// TIA Portal V20 export
FUNCTION_BLOCK "POS3_0_SK_Ablauf"   // FB26, GRAPH
// stored: GraphVersion 6.0, InitialValuesAcquisition false, LanguageInNetworks FBD, SetENOAutomatically false
   // inherited from GRAPH_BASE
   VAR_INPUT
      OFF_SQ { ExternalWritable := 'False'} : Bool := false;   // Kette ausschalten
      INIT_SQ { ExternalWritable := 'False'} : Bool := false;   // Kette in Initialzustand versetzen
      ACK_EF { ExternalWritable := 'False'} : Bool := false;   // Alle Fehler und Störungen quittieren
      REG_EF { ExternalWritable := 'False'} : Bool := false;   // Alle Fehler und Störungen registrieren
      ACK_S { ExternalWritable := 'False'} : Bool := false;   // Schritt quittieren, der an Parameter S_NO anliegt
      REG_S { ExternalWritable := 'False'} : Bool := false;   // Schritt registrieren, der an Parameter S_NO anliegt
      HALT_SQ { ExternalWritable := 'False'} : Bool := false;   // Kette sofort anhalten
      HALT_TM { ExternalWritable := 'False'} : Bool := false;   // Zeiten sofort anhalten
      ZERO_OP { ExternalWritable := 'False'} : Bool := false;   // Alle mit N, L, D zugewiesenen Operanden auf 0 setzen
      EN_IL { ExternalWritable := 'False'} : Bool := false;   // Interlockbearbeitung aktivieren
      EN_SV { ExternalWritable := 'False'} : Bool := false;   // Supervisionsbearbeitung aktivieren
      EN_ACKREQ { ExternalWritable := 'False'} : Bool := false;   // Quittierpflicht aktivieren
      EN_SSKIP { ExternalWritable := 'False'} : Bool := false;   // "Schritte überspringen" aktivieren
      DISP_SACT { ExternalWritable := 'False'} : Bool := false;   // Nur aktive Schritte anzeigen
      DISP_SEF { ExternalWritable := 'False'} : Bool := false;   // Nur fehlerhafte und gestörte Schritte anzeigen
      DISP_SALL { ExternalWritable := 'False'} : Bool := false;   // Alle Schritte anzeigen
      S_PREV { ExternalWritable := 'False'} : Bool := false;   // Vorherigen Schritt am Parameter S_NO ausgeben
      S_NEXT { ExternalWritable := 'False'} : Bool := false;   // Nächsten Schritt am Parameter S_NO anzeigen
      SW_AUTO { ExternalWritable := 'False'} : Bool := false;   // Automatischer Betrieb
      SW_TAP { ExternalWritable := 'False'} : Bool := false;   // Halbautomatisch/Weiterschalten mit Transition
      SW_TOP { ExternalWritable := 'False'} : Bool := false;   // Halbautomatisch/Ignoriere Transition
      SW_MAN { ExternalWritable := 'False'} : Bool := false;   // Handbetrieb
      S_SEL { ExternalWritable := 'False'} : Int := 0;   // Schritt auswählen, der an S_NO ausgegeben werden soll
      S_SELOK { ExternalWritable := 'False'} : Bool := false;   // Wert aus S_SEL nach S_NO übernehmen
      S_ON { ExternalWritable := 'False'} : Bool := false;   // Schritt aktivieren, der an Parameter S_NO anliegt
      S_OFF { ExternalWritable := 'False'} : Bool := false;   // Schritt deaktivieren, der an Parameter S_NO anliegt
      T_PREV { ExternalWritable := 'False'} : Bool := false;   // Vorherige Transition an Parameter T_NO anzeigen
      T_NEXT { ExternalWritable := 'False'} : Bool := false;   // Nächste Transition an Parameter T_NO anzeigen
      T_PUSH { ExternalWritable := 'False'} : Bool := false;   // Schaltfreigabe für Transition im halbautomatischen Betrieb
      EN_LMODE { ExternalWritable := 'False'} : Bool := false;   // Lernmodus aktivieren
   END_VAR
   VAR_OUTPUT
      S_NO { ExternalWritable := 'False'} : Int := 0;   // Schrittnummer
      S_MORE { ExternalWritable := 'False'} : Bool := false;   // Weitere Schritte sind vorhanden und können in S_NO angezeigt werden.
      S_ACTIVE { ExternalWritable := 'False'} : Bool := false;   // Schritt, der an Parameter S_NO angezeigt wird, ist aktiv
      S_TIME { ExternalWritable := 'False'} : Time := T#0ms;   // Schrittaktivierungszeit
      S_TIMEOK { ExternalWritable := 'False'} : Time := T#0ms;   // Schrittaktivierungszeit fehlerfrei
      S_CRITLOC { ExternalWritable := 'False'} : DWord := 16#0;   // Interlock-Kriterienbits
      S_CRITLOCERR { ExternalWritable := 'False'} : DWord := 16#0;   // Interlock-Kriterienbits bei Ereignis L1
      S_STATE { ExternalWritable := 'False'} : Word := 16#0;   // Schrittzustandsbits
      T_NO { ExternalWritable := 'False'} : Int := 0;   // Transitionsnummer
      T_MORE { ExternalWritable := 'False'} : Bool := false;   // Weitere gültige Transitionen zur Anzeige verfügbar
      T_CRIT { ExternalWritable := 'False'} : DWord := 16#0;   // Transitions-Kriterienbits
      T_CRITOLD { ExternalWritable := 'False'} : DWord := 16#0;   // Transitions-Kriterienbits des letzten Zyklus
      T_CRITFLT { ExternalWritable := 'False'} : DWord := 16#0;   // Transitions-Kriterienbits bei Ereignis V1
      ERROR { ExternalWritable := 'False'} : Bool := false;   // Sammelfehler Interlock
      FAULT { ExternalWritable := 'False'} : Bool := false;   // Sammelfehler Supervision
      ERR_FLT { ExternalWritable := 'False'} : Bool := false;   // Sammelfehler Interlock oder Supervision
      SQ_ISOFF { ExternalWritable := 'False'} : Bool := false;   // Kette ausgeschaltet (kein Schritt aktiv)
      SQ_HALTED { ExternalWritable := 'False'} : Bool := false;   // Kette angehalten
      TM_HALTED { ExternalWritable := 'False'} : Bool := false;   // Zeiten angehalten
      OP_ZEROED { ExternalWritable := 'False'} : Bool := false;   // Alle mit N, L oder D zugewiesenen Operanden auf 0 gesetzt
      IL_ENABLED { ExternalWritable := 'False'} : Bool := false;   // Interlockbearbeitung aktiv
      SV_ENABLED { ExternalWritable := 'False'} : Bool := false;   // Supervisionsbearbeitung aktiviert
      ACKREQ_ENABLED { ExternalWritable := 'False'} : Bool := false;   // Quittierpflicht aktiviert
      SSKIP_ENABLED { ExternalWritable := 'False'} : Bool := false;   // Schritte überspringen aktiviert
      SACT_DISP { ExternalWritable := 'False'} : Bool := false;   // Nur aktive Schritte anzeigen
      SEF_DISP { ExternalWritable := 'False'} : Bool := false;   // Nur fehlerhafte oder gestörte Schritte anzeigen
      SALL_DISP { ExternalWritable := 'False'} : Bool := false;   // Alle Schritte anzeigen
      AUTO_ON { ExternalWritable := 'False'} : Bool := false;   // Automatischer Betrieb eingeschaltet
      TAP_ON { ExternalWritable := 'False'} : Bool := false;   // Halbautomatischer Betrieb/Schritt mit Transition eingeschaltet
      TOP_ON { ExternalWritable := 'False'} : Bool := false;   // Halbautomatischer Betrieb/Ignoriere Transition eingeschaltet
      MAN_ON { ExternalWritable := 'False'} : Bool := false;   // Handbetrieb eingeschaltet
      LMODE_ENABLED { ExternalWritable := 'False'} : Bool := false;   // Lernmodus aktiv
   END_VAR
BEGIN
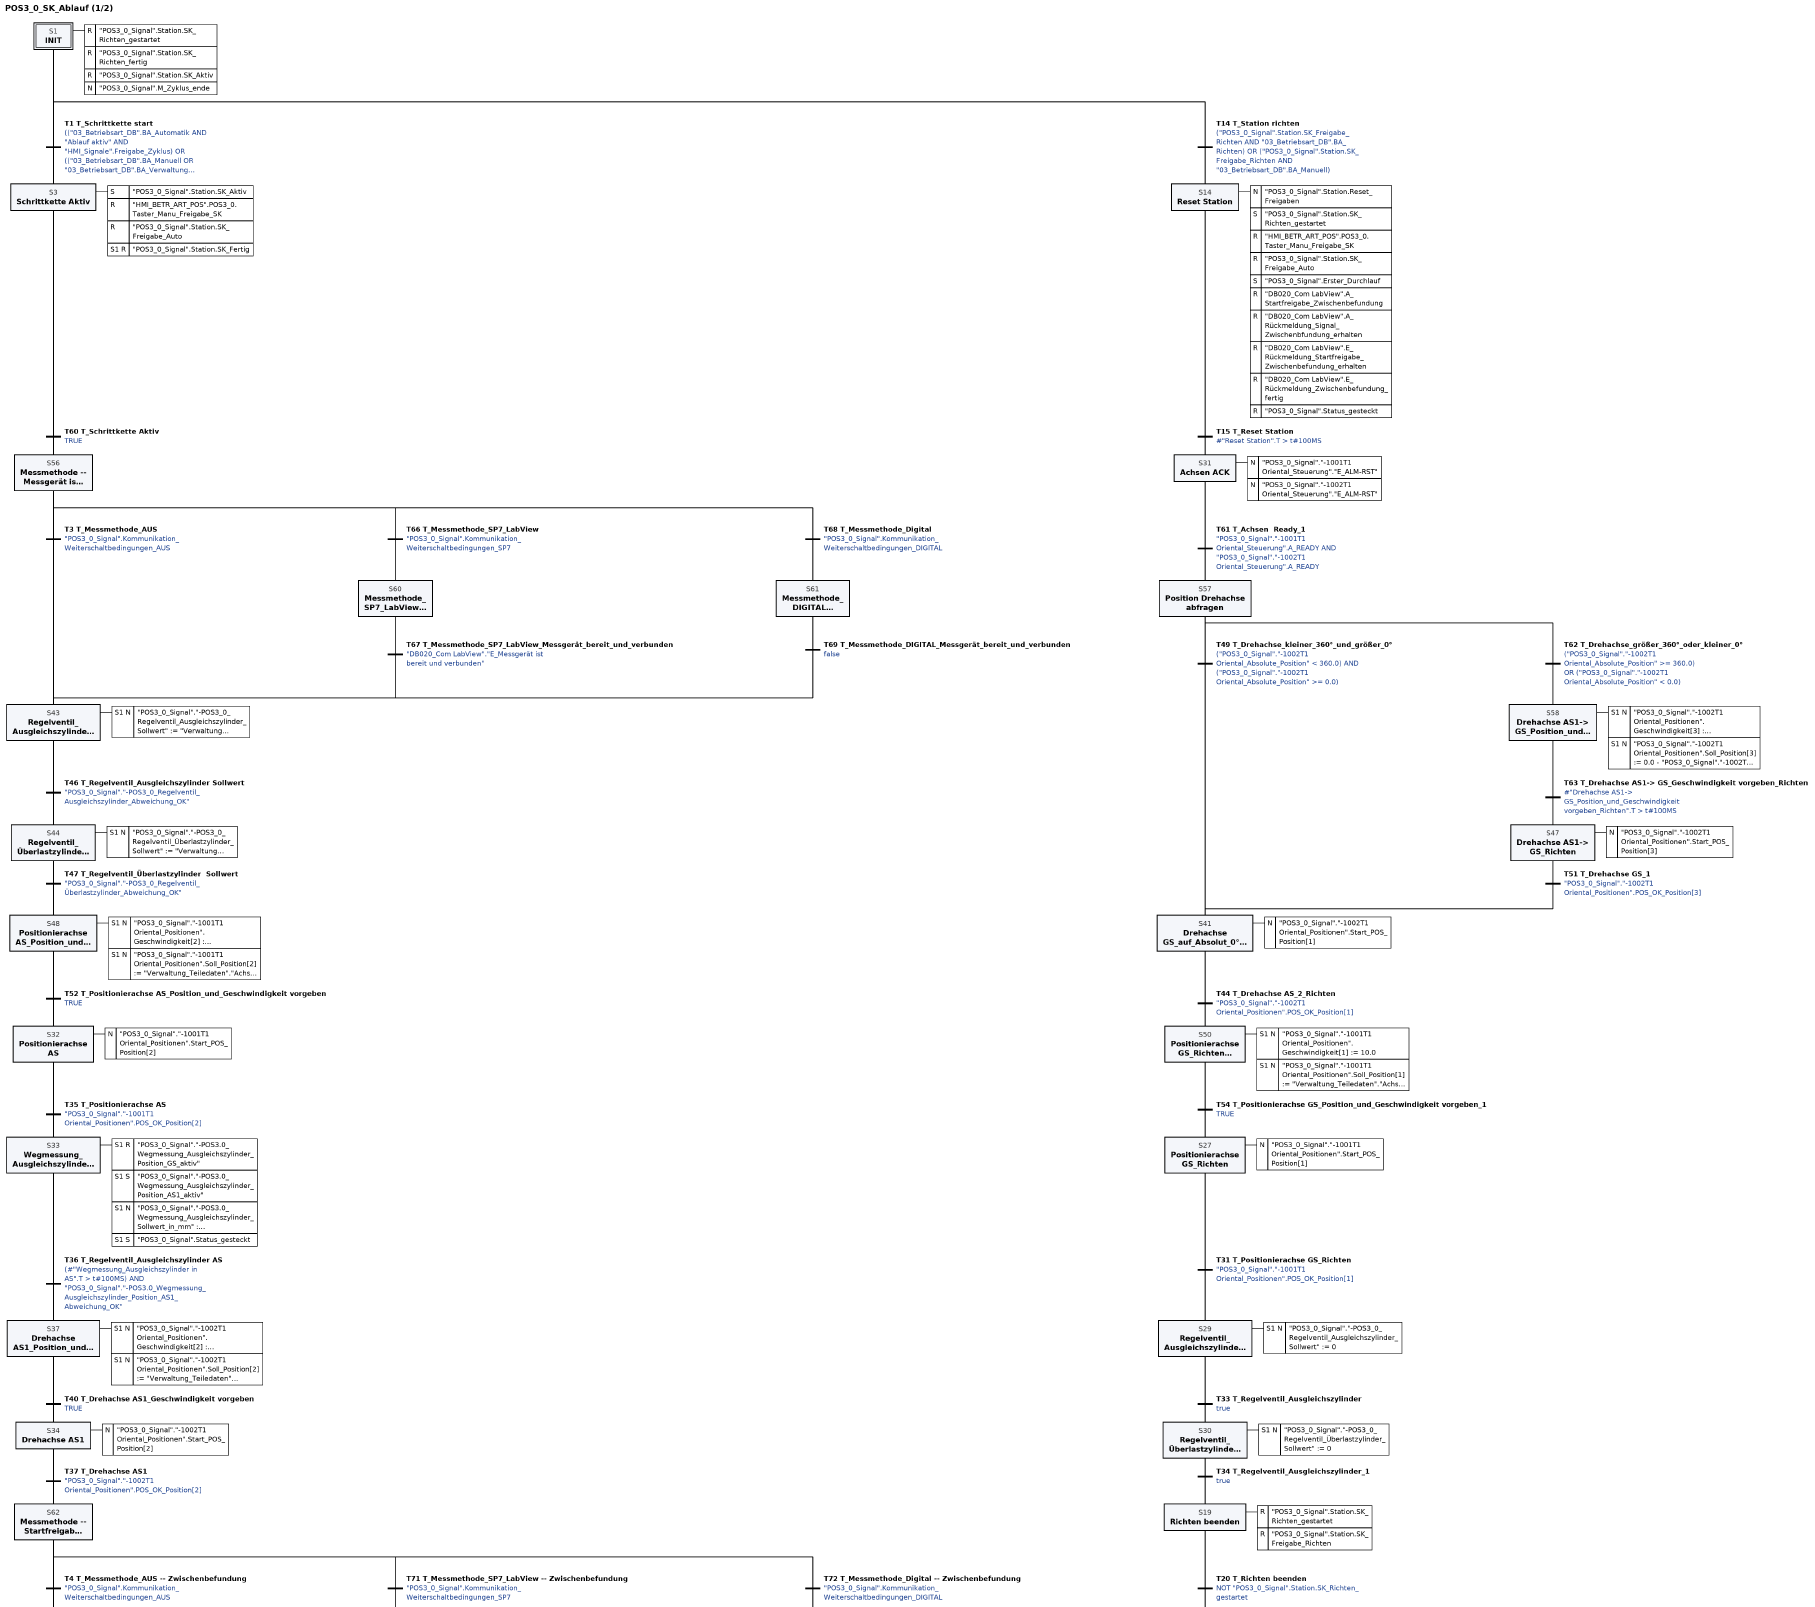
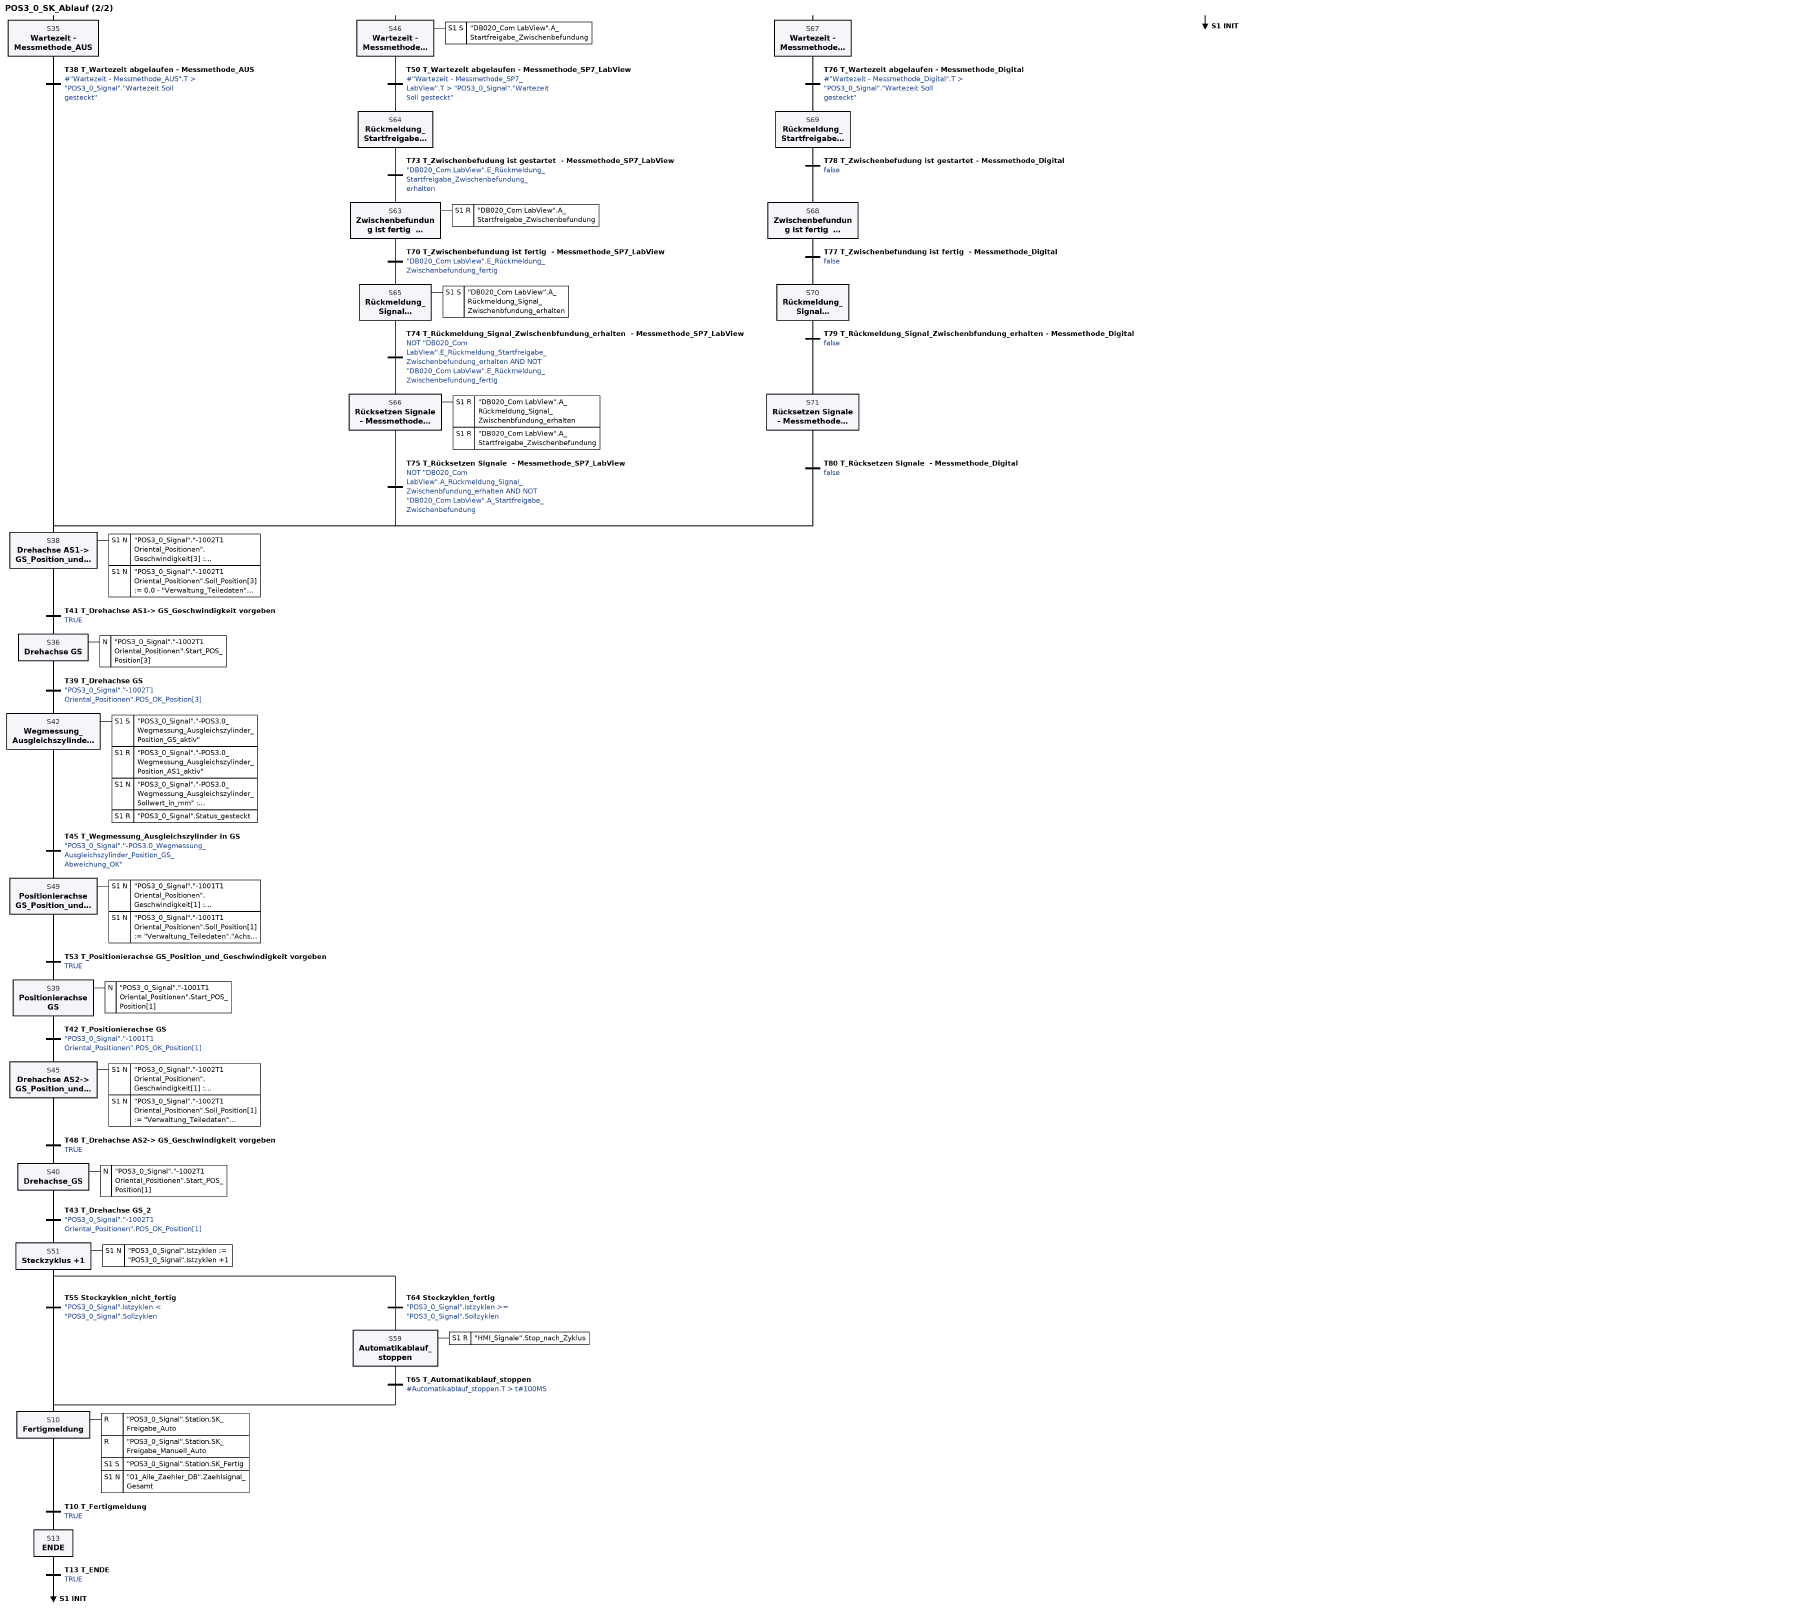
   // sequencer 1
   INITIAL_STEP INIT:   // S1, max time T#10S, warning time T#7S
              R    "POS3_0_Signal".Station.SK_Richten_gestartet
              R    "POS3_0_Signal".Station.SK_Richten_fertig
              R    "POS3_0_Signal".Station.SK_Aktiv
              N    "POS3_0_Signal".M_Zyklus_ende
   END_STEP
   TRANSITION "T_Schrittkette start" FROM INIT TO "Schrittkette Aktiv"   // T1
      := (("03_Betriebsart_DB".BA_Automatik AND "Ablauf aktiv" AND "HMI_Signale".Freigabe_Zyklus) OR (("03_Betriebsart_DB".BA_Manuell OR "03_Betriebsart_DB".BA_Verwaltung) AND "HMI_BETR_ART_POS".POS3_0.Taster_Manu_Freigabe_SK)) AND "Global_Signal"."M_Grundstellung_POS3.0";
   END_TRANSITION
   TRANSITION "T_Station richten" FROM INIT TO "Reset Station"   // T14
      := ("POS3_0_Signal".Station.SK_Freigabe_Richten AND "03_Betriebsart_DB".BA_Richten) OR ("POS3_0_Signal".Station.SK_Freigabe_Richten AND "03_Betriebsart_DB".BA_Manuell);
   END_TRANSITION
   STEP "Schrittkette Aktiv":   // S3, max time T#10S, warning time T#7S
      supervision V := #"Schrittkette Aktiv".U > #"Schrittkette Aktiv".T_MAX;
              S    "POS3_0_Signal".Station.SK_Aktiv
              R    "HMI_BETR_ART_POS".POS3_0.Taster_Manu_Freigabe_SK
              R    "POS3_0_Signal".Station.SK_Freigabe_Auto
          S1  R    "POS3_0_Signal".Station.SK_Fertig
   END_STEP
   TRANSITION "T_Schrittkette Aktiv" FROM "Schrittkette Aktiv" TO "Messmethode -- Messgerät ist bereit oder nicht verbunden"   // T60
      := TRUE;
   END_TRANSITION
   STEP "Drehachse GS":   // S36, max time T#10S, warning time T#7S
      supervision V := #"Drehachse GS".U > #"Drehachse GS".T_MAX;
              N    "POS3_0_Signal"."-1002T1 Oriental_Positionen".Start_POS_Position[3]
   END_STEP
   TRANSITION "T_Drehachse GS" FROM "Drehachse GS" TO "Wegmessung_Ausgleichszylinder in GS"   // T39
      := "POS3_0_Signal"."-1002T1 Oriental_Positionen".POS_OK_Position[3];
   END_TRANSITION
   STEP Fertigmeldung:   // S10, max time T#10S, warning time T#7S
      supervision V := #Fertigmeldung.U > #Fertigmeldung.T_MAX;
              R    "POS3_0_Signal".Station.SK_Freigabe_Auto
              R    "POS3_0_Signal".Station.SK_Freigabe_Manuell_Auto
          S1  S    "POS3_0_Signal".Station.SK_Fertig
          S1  N    "01_Alle_Zaehler_DB".Zaehlsignal_Gesamt
   END_STEP
   TRANSITION T_Fertigmeldung FROM Fertigmeldung TO ENDE   // T10
      := TRUE;
   END_TRANSITION
   STEP ENDE:   // S13, max time T#10S, warning time T#7S
   END_STEP
   TRANSITION T_ENDE FROM ENDE TO INIT   // T13, jump
      := TRUE;
   END_TRANSITION
   STEP "Reset Station":   // S14, max time T#10S, warning time T#7S
              N    "POS3_0_Signal".Station.Reset_Freigaben
              S    "POS3_0_Signal".Station.SK_Richten_gestartet
              R    "HMI_BETR_ART_POS".POS3_0.Taster_Manu_Freigabe_SK
              R    "POS3_0_Signal".Station.SK_Freigabe_Auto
              S    "POS3_0_Signal".Erster_Durchlauf
              R    "DB020_Com LabView".A_Startfreigabe_Zwischenbefundung
              R    "DB020_Com LabView".A_Rückmeldung_Signal_Zwischenbfundung_erhalten
              R    "DB020_Com LabView".E_Rückmeldung_Startfreigabe_Zwischenbefundung_erhalten
              R    "DB020_Com LabView".E_Rückmeldung_Zwischenbefundung_fertig
              R    "POS3_0_Signal".Status_gesteckt
   END_STEP
   TRANSITION "T_Reset Station" FROM "Reset Station" TO "Achsen ACK"   // T15
      := #"Reset Station".T > t#100MS;
   END_TRANSITION
   STEP "Richten beenden":   // S19, max time T#10S, warning time T#7S
              R    "POS3_0_Signal".Station.SK_Richten_gestartet
              R    "POS3_0_Signal".Station.SK_Freigabe_Richten
   END_STEP
   TRANSITION "T_Richten beenden" FROM "Richten beenden" TO INIT   // T20, jump
      := NOT "POS3_0_Signal".Station.SK_Richten_gestartet;
   END_TRANSITION
   STEP "Wartezeit - Messmethode_AUS":   // S35, max time T#10S, warning time T#7S
   END_STEP
   TRANSITION "T_Wartezeit abgelaufen - Messmethode_AUS" FROM "Wartezeit - Messmethode_AUS" TO "Drehachse AS1-> GS_Position_und_Geschwindigkeit vorgeben"   // T38
      := #"Wartezeit - Messmethode_AUS".T > "POS3_0_Signal"."Wartezeit Soll gesteckt";
   END_TRANSITION
   STEP "Positionierachse GS_Richten":   // S27, max time T#10S, warning time T#7S
      supervision V := #"Positionierachse GS_Richten".U > #"Positionierachse GS_Richten".T_MAX;
              N    "POS3_0_Signal"."-1001T1 Oriental_Positionen".Start_POS_Position[1]
   END_STEP
   TRANSITION "T_Positionierachse GS_Richten" FROM "Positionierachse GS_Richten" TO "Regelventil_Ausgleichszylinder auf 0 mbar"   // T31
      := "POS3_0_Signal"."-1001T1 Oriental_Positionen".POS_OK_Position[1];
   END_TRANSITION
   STEP "Achsen ACK":   // S31, max time T#10S, warning time T#7S
              N    "POS3_0_Signal"."-1001T1 Oriental_Steuerung"."E_ALM-RST"
              N    "POS3_0_Signal"."-1002T1 Oriental_Steuerung"."E_ALM-RST"
   END_STEP
   TRANSITION "T_Achsen  Ready_1" FROM "Achsen ACK" TO "Position Drehachse abfragen"   // T61
      := "POS3_0_Signal"."-1001T1 Oriental_Steuerung".A_READY AND "POS3_0_Signal"."-1002T1 Oriental_Steuerung".A_READY;
   END_TRANSITION
   STEP "Regelventil_Ausgleichszylinder auf 0 mbar":   // S29, max time T#10S, warning time T#7S
          S1  N    "POS3_0_Signal"."-POS3_0_Regelventil_Ausgleichszylinder_Sollwert" := 0
   END_STEP
   TRANSITION T_Regelventil_Ausgleichszylinder FROM "Regelventil_Ausgleichszylinder auf 0 mbar" TO "Regelventil_Überlastzylinder auf 0 mbar"   // T33
      := true;
   END_TRANSITION
   STEP "Regelventil_Überlastzylinder auf 0 mbar":   // S30, max time T#10S, warning time T#7S
          S1  N    "POS3_0_Signal"."-POS3_0_Regelventil_Überlastzylinder_Sollwert" := 0
   END_STEP
   TRANSITION T_Regelventil_Ausgleichszylinder_1 FROM "Regelventil_Überlastzylinder auf 0 mbar" TO "Richten beenden"   // T34
      := true;
   END_TRANSITION
   STEP "Positionierachse AS":   // S32, max time T#10S, warning time T#7S
      supervision V := #"Positionierachse AS".U > t#300s;
              N    "POS3_0_Signal"."-1001T1 Oriental_Positionen".Start_POS_Position[2]
   END_STEP
   TRANSITION "T_Positionierachse AS" FROM "Positionierachse AS" TO "Wegmessung_Ausgleichszylinder in AS"   // T35
      := "POS3_0_Signal"."-1001T1 Oriental_Positionen".POS_OK_Position[2];
   END_TRANSITION
   STEP "Wegmessung_Ausgleichszylinder in AS":   // S33, max time T#10S, warning time T#7S
      supervision V := #"Wegmessung_Ausgleichszylinder in AS".U > #"Wegmessung_Ausgleichszylinder in AS".T_MAX;
          S1  R    "POS3_0_Signal"."-POS3.0_Wegmessung_Ausgleichszylinder_Position_GS_aktiv"
          S1  S    "POS3_0_Signal"."-POS3.0_Wegmessung_Ausgleichszylinder_Position_AS1_aktiv"
          S1  N    "POS3_0_Signal"."-POS3.0_Wegmessung_Ausgleichszylinder_Sollwert_in_mm" := "Verwaltung_Teiledaten"."Wegmessung_Ausgleichszylinder Position AS1"
          S1  S    "POS3_0_Signal".Status_gesteckt
   END_STEP
   TRANSITION "T_Regelventil_Ausgleichszylinder AS" FROM "Wegmessung_Ausgleichszylinder in AS" TO "Drehachse AS1_Position_und_Geschwindigkeit vorgeben"   // T36
      := (#"Wegmessung_Ausgleichszylinder in AS".T > t#100MS) AND "POS3_0_Signal"."-POS3.0_Wegmessung_Ausgleichszylinder_Position_AS1_Abweichung_OK";
   END_TRANSITION
   STEP "Drehachse AS1":   // S34, max time T#10S, warning time T#7S
      supervision V := #"Drehachse AS1".U > #"Drehachse AS1".T_MAX;
              N    "POS3_0_Signal"."-1002T1 Oriental_Positionen".Start_POS_Position[2]
   END_STEP
   TRANSITION "T_Drehachse AS1" FROM "Drehachse AS1" TO "Messmethode -- Startfreigabe Zwischenbefundung"   // T37
      := "POS3_0_Signal"."-1002T1 Oriental_Positionen".POS_OK_Position[2];
   END_TRANSITION
   STEP "Positionierachse GS":   // S39, max time T#10S, warning time T#7S
      supervision V := #"Positionierachse GS".U > t#300s;
              N    "POS3_0_Signal"."-1001T1 Oriental_Positionen".Start_POS_Position[1]
   END_STEP
   TRANSITION "T_Positionierachse GS" FROM "Positionierachse GS" TO "Drehachse AS2-> GS_Position_und_Geschwindigkeit vorgeben"   // T42
      := "POS3_0_Signal"."-1001T1 Oriental_Positionen".POS_OK_Position[1];
   END_TRANSITION
   STEP Drehachse_GS:   // S40, max time T#10S, warning time T#7S
      supervision V := #Drehachse_GS.U > #Drehachse_GS.T_MAX;
              N    "POS3_0_Signal"."-1002T1 Oriental_Positionen".Start_POS_Position[1]
   END_STEP
   TRANSITION "T_Drehachse GS_2" FROM Drehachse_GS TO "Steckzyklus +1"   // T43
      := "POS3_0_Signal"."-1002T1 Oriental_Positionen".POS_OK_Position[1];
   END_TRANSITION
   STEP "Drehachse GS_auf_Absolut_0°_Richten":   // S41, max time T#10S, warning time T#7S
      supervision V := #"Drehachse GS_auf_Absolut_0°_Richten".U > #"Drehachse GS_auf_Absolut_0°_Richten".T_MAX;
              N    "POS3_0_Signal"."-1002T1 Oriental_Positionen".Start_POS_Position[1]
   END_STEP
   TRANSITION "T_Drehachse AS_2_Richten" FROM "Drehachse GS_auf_Absolut_0°_Richten" TO "Positionierachse GS_Richten_Position_und_Geschwindigkeit vorgeben"   // T44
      := "POS3_0_Signal"."-1002T1 Oriental_Positionen".POS_OK_Position[1];
   END_TRANSITION
   STEP "Wegmessung_Ausgleichszylinder in GS":   // S42, max time T#10S, warning time T#7S
      supervision V := #"Wegmessung_Ausgleichszylinder in GS".U > #"Wegmessung_Ausgleichszylinder in GS".T_MAX;
          S1  S    "POS3_0_Signal"."-POS3.0_Wegmessung_Ausgleichszylinder_Position_GS_aktiv"
          S1  R    "POS3_0_Signal"."-POS3.0_Wegmessung_Ausgleichszylinder_Position_AS1_aktiv"
          S1  N    "POS3_0_Signal"."-POS3.0_Wegmessung_Ausgleichszylinder_Sollwert_in_mm" := "Verwaltung_Teiledaten"."Wegmessung_Ausgleichszylinder Position GS"
          S1  R    "POS3_0_Signal".Status_gesteckt
   END_STEP
   TRANSITION "T_Wegmessung_Ausgleichszylinder in GS" FROM "Wegmessung_Ausgleichszylinder in GS" TO "Positionierachse GS_Position_und_Geschwindigkeit vorgeben"   // T45
      := "POS3_0_Signal"."-POS3.0_Wegmessung_Ausgleichszylinder_Position_GS_Abweichung_OK";
   END_TRANSITION
   STEP "Regelventil_Überlastzylinder  Sollwert":   // S44, max time T#10S, warning time T#7S
      supervision V := #"Regelventil_Überlastzylinder  Sollwert".U > #"Regelventil_Überlastzylinder  Sollwert".T_MAX;
          S1  N    "POS3_0_Signal"."-POS3_0_Regelventil_Überlastzylinder_Sollwert" := "Verwaltung_Teiledaten"."Druck p2 Überlastzylinder"
   END_STEP
   TRANSITION "T_Regelventil_Überlastzylinder  Sollwert" FROM "Regelventil_Überlastzylinder  Sollwert" TO "Positionierachse AS_Position_und_Geschwindigkeit vorgeben"   // T47
      := "POS3_0_Signal"."-POS3_0_Regelventil_Überlastzylinder_Abweichung_OK";
   END_TRANSITION
   STEP "Drehachse AS1_Position_und_Geschwindigkeit vorgeben":   // S37, max time T#10S, warning time T#7S
      supervision V := #"Drehachse AS1_Position_und_Geschwindigkeit vorgeben".U > #"Drehachse AS1_Position_und_Geschwindigkeit vorgeben".T_MAX;
          S1  N    "POS3_0_Signal"."-1002T1 Oriental_Positionen".Geschwindigkeit[2] := "Verwaltung_Teiledaten"."Drehantrieb Geschwindigkeit GS->AS1" / 6
          S1  N    "POS3_0_Signal"."-1002T1 Oriental_Positionen".Soll_Position[2] := "Verwaltung_Teiledaten"."Drehantrieb Position AS1"
   END_STEP
   TRANSITION "T_Drehachse AS1_Geschwindigkeit vorgeben" FROM "Drehachse AS1_Position_und_Geschwindigkeit vorgeben" TO "Drehachse AS1"   // T40
      := TRUE;
   END_TRANSITION
   STEP "Drehachse AS1-> GS_Position_und_Geschwindigkeit vorgeben":   // S38, max time T#10S, warning time T#7S
      supervision V := #"Drehachse AS1-> GS_Position_und_Geschwindigkeit vorgeben".U > #"Drehachse AS1-> GS_Position_und_Geschwindigkeit vorgeben".T_MAX;
          S1  N    "POS3_0_Signal"."-1002T1 Oriental_Positionen".Geschwindigkeit[3] := "Verwaltung_Teiledaten"."Drehantrieb Geschwindigkeit AS1->GS" / 6
          S1  N    "POS3_0_Signal"."-1002T1 Oriental_Positionen".Soll_Position[3] := 0.0 - "Verwaltung_Teiledaten"."Drehantrieb Position AS1"
   END_STEP
   TRANSITION "T_Drehachse AS1-> GS_Geschwindigkeit vorgeben" FROM "Drehachse AS1-> GS_Position_und_Geschwindigkeit vorgeben" TO "Drehachse GS"   // T41
      := TRUE;
   END_TRANSITION
   STEP "Regelventil_Ausgleichszylinder Sollwert":   // S43, max time T#10S, warning time T#7S
      supervision V := #"Regelventil_Ausgleichszylinder Sollwert".U > #"Regelventil_Ausgleichszylinder Sollwert".T_MAX;
          S1  N    "POS3_0_Signal"."-POS3_0_Regelventil_Ausgleichszylinder_Sollwert" := "Verwaltung_Teiledaten"."Druck p1 Ausgleichszylinder"
   END_STEP
   TRANSITION "T_Regelventil_Ausgleichszylinder Sollwert" FROM "Regelventil_Ausgleichszylinder Sollwert" TO "Regelventil_Überlastzylinder  Sollwert"   // T46
      := "POS3_0_Signal"."-POS3_0_Regelventil_Ausgleichszylinder_Abweichung_OK";
   END_TRANSITION
   STEP "Drehachse AS2-> GS_Position_und_Geschwindigkeit vorgeben":   // S45, max time T#10S, warning time T#7S
      supervision V := #"Drehachse AS2-> GS_Position_und_Geschwindigkeit vorgeben".U > #"Drehachse AS2-> GS_Position_und_Geschwindigkeit vorgeben".T_MAX;
          S1  N    "POS3_0_Signal"."-1002T1 Oriental_Positionen".Geschwindigkeit[1] := "Verwaltung_Teiledaten"."Drehantrieb Motorstrombegrenzung" / 6
          S1  N    "POS3_0_Signal"."-1002T1 Oriental_Positionen".Soll_Position[1] := "Verwaltung_Teiledaten"."Drehantrieb Position GS"
   END_STEP
   TRANSITION "T_Drehachse AS2-> GS_Geschwindigkeit vorgeben" FROM "Drehachse AS2-> GS_Position_und_Geschwindigkeit vorgeben" TO Drehachse_GS   // T48
      := TRUE;
   END_TRANSITION
   STEP "Positionierachse AS_Position_und_Geschwindigkeit vorgeben":   // S48, max time T#10S, warning time T#7S
      supervision V := #"Positionierachse AS_Position_und_Geschwindigkeit vorgeben".U > #"Positionierachse AS_Position_und_Geschwindigkeit vorgeben".T_MAX;
          S1  N    "POS3_0_Signal"."-1001T1 Oriental_Positionen".Geschwindigkeit[2] := "Verwaltung_Teiledaten"."Achse Geschwindigkeit GS->AS" / 150
          S1  N    "POS3_0_Signal"."-1001T1 Oriental_Positionen".Soll_Position[2] := "Verwaltung_Teiledaten"."Achse Position AS"
   END_STEP
   TRANSITION "T_Positionierachse AS_Position_und_Geschwindigkeit vorgeben" FROM "Positionierachse AS_Position_und_Geschwindigkeit vorgeben" TO "Positionierachse AS"   // T52
      := TRUE;
   END_TRANSITION
   STEP "Positionierachse GS_Position_und_Geschwindigkeit vorgeben":   // S49, max time T#10S, warning time T#7S
      supervision V := #"Positionierachse GS_Position_und_Geschwindigkeit vorgeben".U > #"Positionierachse GS_Position_und_Geschwindigkeit vorgeben".T_MAX;
          S1  N    "POS3_0_Signal"."-1001T1 Oriental_Positionen".Geschwindigkeit[1] := "Verwaltung_Teiledaten"."Achse Geschwindigkeit AS->GS" / 150
          S1  N    "POS3_0_Signal"."-1001T1 Oriental_Positionen".Soll_Position[1] := "Verwaltung_Teiledaten"."Achse Position GS"
   END_STEP
   TRANSITION "T_Positionierachse GS_Position_und_Geschwindigkeit vorgeben" FROM "Positionierachse GS_Position_und_Geschwindigkeit vorgeben" TO "Positionierachse GS"   // T53
      := TRUE;
   END_TRANSITION
   STEP "Positionierachse GS_Richten_Position_und_Geschwindigkeit vorgeben":   // S50, max time T#10S, warning time T#7S
      supervision V := #"Positionierachse GS_Richten_Position_und_Geschwindigkeit vorgeben".U > #"Positionierachse GS_Richten_Position_und_Geschwindigkeit vorgeben".T_MAX;
          S1  N    "POS3_0_Signal"."-1001T1 Oriental_Positionen".Geschwindigkeit[1] := 10.0
          S1  N    "POS3_0_Signal"."-1001T1 Oriental_Positionen".Soll_Position[1] := "Verwaltung_Teiledaten"."Achse Position GS"
   END_STEP
   TRANSITION "T_Positionierachse GS_Position_und_Geschwindigkeit vorgeben_1" FROM "Positionierachse GS_Richten_Position_und_Geschwindigkeit vorgeben" TO "Positionierachse GS_Richten"   // T54
      := TRUE;
   END_TRANSITION
   STEP "Steckzyklus +1":   // S51, max time T#10S, warning time T#7S
          S1  N    "POS3_0_Signal".Istzyklen := "POS3_0_Signal".Istzyklen +1
   END_STEP
   TRANSITION Steckzyklen_nicht_fertig FROM "Steckzyklus +1" TO Fertigmeldung   // T55
      := "POS3_0_Signal".Istzyklen < "POS3_0_Signal".Sollzyklen;
   END_TRANSITION
   TRANSITION Steckzyklen_fertig FROM "Steckzyklus +1" TO Automatikablauf_stoppen   // T64
      := "POS3_0_Signal".Istzyklen >= "POS3_0_Signal".Sollzyklen;
   END_TRANSITION
   STEP "Messmethode -- Messgerät ist bereit oder nicht verbunden":   // S56, max time T#10S, warning time T#7S
      supervision V := #"Messmethode -- Messgerät ist bereit oder nicht verbunden".U > T#30s;
   END_STEP
   TRANSITION T_Messmethode_AUS FROM "Messmethode -- Messgerät ist bereit oder nicht verbunden" TO "Regelventil_Ausgleichszylinder Sollwert"   // T3
      := "POS3_0_Signal".Kommunikation_Weiterschaltbedingungen_AUS;
   END_TRANSITION
   TRANSITION T_Messmethode_SP7_LabView FROM "Messmethode -- Messgerät ist bereit oder nicht verbunden" TO Messmethode_SP7_LabView_Messgerät_bereit_und_verbunden   // T66
      := "POS3_0_Signal".Kommunikation_Weiterschaltbedingungen_SP7;
   END_TRANSITION
   TRANSITION T_Messmethode_Digital FROM "Messmethode -- Messgerät ist bereit oder nicht verbunden" TO Messmethode_DIGITAL_Messgerät_bereit_und_verbunden   // T68
      := "POS3_0_Signal".Kommunikation_Weiterschaltbedingungen_DIGITAL;
   END_TRANSITION
   STEP "Position Drehachse abfragen":   // S57, max time T#10S, warning time T#7S
   END_STEP
   TRANSITION "T_Drehachse_kleiner_360°_und_größer_0°" FROM "Position Drehachse abfragen" TO "Drehachse GS_auf_Absolut_0°_Richten"   // T49
      := ("POS3_0_Signal"."-1002T1 Oriental_Absolute_Position" < 360.0) AND ("POS3_0_Signal"."-1002T1 Oriental_Absolute_Position" >= 0.0);
   END_TRANSITION
   TRANSITION "T_Drehachse_größer_360°_oder_kleiner_0°" FROM "Position Drehachse abfragen" TO "Drehachse AS1-> GS_Position_und_Geschwindigkeit vorgeben_Richten"   // T62
      := ("POS3_0_Signal"."-1002T1 Oriental_Absolute_Position" >= 360.0) OR ("POS3_0_Signal"."-1002T1 Oriental_Absolute_Position" < 0.0);
   END_TRANSITION
   STEP "Drehachse AS1-> GS_Richten":   // S47, max time T#10S, warning time T#7S
      supervision V := #"Drehachse AS1-> GS_Richten".U > #"Drehachse AS1-> GS_Richten".T_MAX;
              N    "POS3_0_Signal"."-1002T1 Oriental_Positionen".Start_POS_Position[3]
   END_STEP
   TRANSITION "T_Drehachse GS_1" FROM "Drehachse AS1-> GS_Richten" TO "Drehachse GS_auf_Absolut_0°_Richten"   // T51
      := "POS3_0_Signal"."-1002T1 Oriental_Positionen".POS_OK_Position[3];
   END_TRANSITION
   STEP "Drehachse AS1-> GS_Position_und_Geschwindigkeit vorgeben_Richten":   // S58, max time T#10S, warning time T#7S
      supervision V := #"Drehachse AS1-> GS_Position_und_Geschwindigkeit vorgeben_Richten".U > #"Drehachse AS1-> GS_Position_und_Geschwindigkeit vorgeben_Richten".T_MAX;
          S1  N    "POS3_0_Signal"."-1002T1 Oriental_Positionen".Geschwindigkeit[3] := "Verwaltung_Teiledaten"."Drehantrieb Geschwindigkeit AS1->GS" / 6
          S1  N    "POS3_0_Signal"."-1002T1 Oriental_Positionen".Soll_Position[3] := 0.0 - "POS3_0_Signal"."-1002T1 Oriental_Absolute_Position"
   END_STEP
   TRANSITION "T_Drehachse AS1-> GS_Geschwindigkeit vorgeben_Richten" FROM "Drehachse AS1-> GS_Position_und_Geschwindigkeit vorgeben_Richten" TO "Drehachse AS1-> GS_Richten"   // T63
      := #"Drehachse AS1-> GS_Position_und_Geschwindigkeit vorgeben_Richten".T > t#100MS;
   END_TRANSITION
   STEP Automatikablauf_stoppen:   // S59, max time T#10S, warning time T#7S
          S1  R    "HMI_Signale".Stop_nach_Zyklus
   END_STEP
   TRANSITION T_Automatikablauf_stoppen FROM Automatikablauf_stoppen TO Fertigmeldung   // T65
      := #Automatikablauf_stoppen.T > t#100MS;
   END_TRANSITION
   STEP Messmethode_SP7_LabView_Messgerät_bereit_und_verbunden:   // S60, max time T#10S, warning time T#7S
   END_STEP
   TRANSITION T_Messmethode_SP7_LabView_Messgerät_bereit_und_verbunden FROM Messmethode_SP7_LabView_Messgerät_bereit_und_verbunden TO "Regelventil_Ausgleichszylinder Sollwert"   // T67
      := "DB020_Com LabView"."E_Messgerät ist bereit und verbunden";
   END_TRANSITION
   STEP Messmethode_DIGITAL_Messgerät_bereit_und_verbunden:   // S61, max time T#10S, warning time T#7S
   END_STEP
   TRANSITION T_Messmethode_DIGITAL_Messgerät_bereit_und_verbunden FROM Messmethode_DIGITAL_Messgerät_bereit_und_verbunden TO "Regelventil_Ausgleichszylinder Sollwert"   // T69
      := false;
   END_TRANSITION
   STEP "Messmethode -- Startfreigabe Zwischenbefundung":   // S62, max time T#10S, warning time T#7S
   END_STEP
   TRANSITION "T_Messmethode_AUS -- Zwischenbefundung" FROM "Messmethode -- Startfreigabe Zwischenbefundung" TO "Wartezeit - Messmethode_AUS"   // T4
      := "POS3_0_Signal".Kommunikation_Weiterschaltbedingungen_AUS;
   END_TRANSITION
   TRANSITION "T_Messmethode_SP7_LabView -- Zwischenbefundung" FROM "Messmethode -- Startfreigabe Zwischenbefundung" TO "Wartezeit - Messmethode_SP7_LabView"   // T71
      := "POS3_0_Signal".Kommunikation_Weiterschaltbedingungen_SP7;
   END_TRANSITION
   TRANSITION "T_Messmethode_Digital -- Zwischenbefundung" FROM "Messmethode -- Startfreigabe Zwischenbefundung" TO "Wartezeit - Messmethode_Digital"   // T72
      := "POS3_0_Signal".Kommunikation_Weiterschaltbedingungen_DIGITAL;
   END_TRANSITION
   STEP "Wartezeit - Messmethode_SP7_LabView":   // S46, max time T#10S, warning time T#7S
          S1  S    "DB020_Com LabView".A_Startfreigabe_Zwischenbefundung
   END_STEP
   TRANSITION "T_Wartezeit abgelaufen - Messmethode_SP7_LabView" FROM "Wartezeit - Messmethode_SP7_LabView" TO "Rückmeldung_Startfreigabe_Zwischenbefundung_erhalten - Messmethode_SP7_LabView"   // T50
      := #"Wartezeit - Messmethode_SP7_LabView".T > "POS3_0_Signal"."Wartezeit Soll gesteckt";
   END_TRANSITION
   STEP "Zwischenbefundung ist fertig  - Messmethode_SP7_LabView":   // S63, max time T#10S, warning time T#7S
      supervision V := #"Zwischenbefundung ist fertig  - Messmethode_SP7_LabView".U > T#30s;
          S1  R    "DB020_Com LabView".A_Startfreigabe_Zwischenbefundung
   END_STEP
   TRANSITION "T_Zwischenbefundung ist fertig  - Messmethode_SP7_LabView" FROM "Zwischenbefundung ist fertig  - Messmethode_SP7_LabView" TO "Rückmeldung_Signal_Zwischenbfundung_erhalten  - Messmethode_SP7_LabView"   // T70
      := "DB020_Com LabView".E_Rückmeldung_Zwischenbefundung_fertig;
   END_TRANSITION
   STEP "Rückmeldung_Startfreigabe_Zwischenbefundung_erhalten - Messmethode_SP7_LabView":   // S64, max time T#10S, warning time T#7S
      supervision V := #"Rückmeldung_Startfreigabe_Zwischenbefundung_erhalten - Messmethode_SP7_LabView".U > t#30s;
   END_STEP
   TRANSITION "T_Zwischenbefudung ist gestartet  - Messmethode_SP7_LabView" FROM "Rückmeldung_Startfreigabe_Zwischenbefundung_erhalten - Messmethode_SP7_LabView" TO "Zwischenbefundung ist fertig  - Messmethode_SP7_LabView"   // T73
      := "DB020_Com LabView".E_Rückmeldung_Startfreigabe_Zwischenbefundung_erhalten;
   END_TRANSITION
   STEP "Rückmeldung_Signal_Zwischenbfundung_erhalten  - Messmethode_SP7_LabView":   // S65, max time T#10S, warning time T#7S
      supervision V := #"Rückmeldung_Signal_Zwischenbfundung_erhalten  - Messmethode_SP7_LabView".U > t#30S;
          S1  S    "DB020_Com LabView".A_Rückmeldung_Signal_Zwischenbfundung_erhalten
   END_STEP
   TRANSITION "T_Rückmeldung_Signal_Zwischenbfundung_erhalten  - Messmethode_SP7_LabView" FROM "Rückmeldung_Signal_Zwischenbfundung_erhalten  - Messmethode_SP7_LabView" TO "Rücksetzen Signale  - Messmethode_SP7_LabView"   // T74
      := NOT "DB020_Com LabView".E_Rückmeldung_Startfreigabe_Zwischenbefundung_erhalten AND NOT "DB020_Com LabView".E_Rückmeldung_Zwischenbefundung_fertig;
   END_TRANSITION
   STEP "Rücksetzen Signale  - Messmethode_SP7_LabView":   // S66, max time T#10S, warning time T#7S
      supervision V := #"Rücksetzen Signale  - Messmethode_SP7_LabView".U > t#30S;
          S1  R    "DB020_Com LabView".A_Rückmeldung_Signal_Zwischenbfundung_erhalten
          S1  R    "DB020_Com LabView".A_Startfreigabe_Zwischenbefundung
   END_STEP
   TRANSITION "T_Rücksetzen Signale  - Messmethode_SP7_LabView" FROM "Rücksetzen Signale  - Messmethode_SP7_LabView" TO "Drehachse AS1-> GS_Position_und_Geschwindigkeit vorgeben"   // T75
      := NOT "DB020_Com LabView".A_Rückmeldung_Signal_Zwischenbfundung_erhalten AND NOT "DB020_Com LabView".A_Startfreigabe_Zwischenbefundung;
   END_TRANSITION
   STEP "Wartezeit - Messmethode_Digital":   // S67, max time T#10S, warning time T#7S
   END_STEP
   TRANSITION "T_Wartezeit abgelaufen - Messmethode_Digital" FROM "Wartezeit - Messmethode_Digital" TO "Rückmeldung_Startfreigabe_Zwischenbefundung_erhalten - Messmethode_Digital"   // T76
      := #"Wartezeit - Messmethode_Digital".T > "POS3_0_Signal"."Wartezeit Soll gesteckt";
   END_TRANSITION
   STEP "Zwischenbefundung ist fertig  - Messmethode_Digital":   // S68, max time T#10S, warning time T#7S
      supervision V := #"Zwischenbefundung ist fertig  - Messmethode_Digital".U > T#30s;
   END_STEP
   TRANSITION "T_Zwischenbefundung ist fertig  - Messmethode_Digital" FROM "Zwischenbefundung ist fertig  - Messmethode_Digital" TO "Rückmeldung_Signal_Zwischenbfundung_erhalten - Messmethode_Digital"   // T77
      := false;
   END_TRANSITION
   STEP "Rückmeldung_Startfreigabe_Zwischenbefundung_erhalten - Messmethode_Digital":   // S69, max time T#10S, warning time T#7S
      supervision V := #"Rückmeldung_Startfreigabe_Zwischenbefundung_erhalten - Messmethode_Digital".U > t#30s;
   END_STEP
   TRANSITION "T_Zwischenbefudung ist gestartet - Messmethode_Digital" FROM "Rückmeldung_Startfreigabe_Zwischenbefundung_erhalten - Messmethode_Digital" TO "Zwischenbefundung ist fertig  - Messmethode_Digital"   // T78
      := false;
   END_TRANSITION
   STEP "Rückmeldung_Signal_Zwischenbfundung_erhalten - Messmethode_Digital":   // S70, max time T#10S, warning time T#7S
      supervision V := #"Rückmeldung_Signal_Zwischenbfundung_erhalten - Messmethode_Digital".U > t#30S;
   END_STEP
   TRANSITION "T_Rückmeldung_Signal_Zwischenbfundung_erhalten - Messmethode_Digital" FROM "Rückmeldung_Signal_Zwischenbfundung_erhalten - Messmethode_Digital" TO "Rücksetzen Signale  - Messmethode_Digital"   // T79
      := false;
   END_TRANSITION
   STEP "Rücksetzen Signale  - Messmethode_Digital":   // S71, max time T#10S, warning time T#7S
      supervision V := #"Rücksetzen Signale  - Messmethode_Digital".U > t#30S;
   END_STEP
   TRANSITION "T_Rücksetzen Signale  - Messmethode_Digital" FROM "Rücksetzen Signale  - Messmethode_Digital" TO "Drehachse AS1-> GS_Position_und_Geschwindigkeit vorgeben"   // T80
      := false;
   END_TRANSITION
END_FUNCTION_BLOCK
